FUNCTION F_SpindleClutchStatus : BYTE
(*

The function used to get clutch status.
.0 - Clutch is closed without tool
.1 - Clutch is closed with tool
.2 - Tool is wrong closed in clutch
.3 -  Clutch open and with tool

Constructor: 		Patryk Panylo
Company:		E. Riexinger GmbH
Date:			04.08.2015
Version:			1.00

Date:			Revision:		Who:				Comment
dd.mm.yyyy		x.xx			Initials			comment

*)
VAR_INPUT
	(* Input variables / Eingang Variablen *)
	nClutchStatus 						:INT;						(* AIx.x Status of bit clutch / Spannzange status *)
END_VAR
VAR
	(* Variables *)
	fbScaling						:FB_Scaling;
END_VAR


fbScaling(
	bEnable := TRUE,
	lrInput := INT_TO_LREAL(nClutchStatus),
	lrXLowLimit := 0,
	lrXUpperLimit := 32767,
	lrYLowLimit := 0,
	lrYUpperLimit := 10,
	usiPrecision := 2
);

F_SpindleClutchStatus := 16#0;

IF fbScaling.lrOutputPV >= 5.3
     AND fbScaling.lrOutputPV <= 7.0
THEN
	F_SpindleClutchStatus.0 := TRUE;			(* Clutch is closed without tool *)

ELSIF fbScaling.lrOutputPV >= 3.8
     	    AND fbScaling.lrOutputPV < 5.3
THEN
	F_SpindleClutchStatus.1 := TRUE;			(* Clutch is closed with tool *)

ELSIF fbScaling.lrOutputPV >= 1.4
     	    AND fbScaling.lrOutputPV < 3.8
THEN
	F_SpindleClutchStatus.2 := TRUE;			(* Tool is wrong closed in clutch *)

ELSIF fbScaling.lrOutputPV >= 1.0
     	    AND fbScaling.lrOutputPV < 1.4
THEN
	F_SpindleClutchStatus.3 := TRUE;			(* Clutch without tool *)

END_IF

END_FUNCTION

(* stored: Version 1.1.0.1, ProductVersion 3.1.4024.15
   POU F_SpindleClutchStatus: Id {ea94b708-5a59-4022-9eac-bc8bd1c55ccd}, SpecialFunc None *)
